SUBAPPLICATION Uebung_157 (* Übung zu FsInfo/FsDir: File Server abfragen und Verzeichnis listen *)
  (* Standard: 61499-2; Description: Copyright (c) 2026 Meisterschulen am Ostbahnhof This program and the accompanying materials are made available under the terms of the Eclipse Public License 2.0 which is available at https://www.eclipse.org/legal/epl-2.0/ SPDX-License-Identifier: EPL-2.0 *)
  (* Version 1.0, 2026-11-26, Franz Höpfinger, Meisterschulen am Ostbahnhof, initial API and implementation and/or initial documentation *)
  PACKAGE Uebungen;
  IMPORT Uebungen::const::Uebung_150_159::FileServer::FS_ADD;
  IMPORT Uebungen::const::Uebung_150_159::FileServer::FS_FLT;
  IMPORT Uebungen::const::Uebung_150_159::FileServer::FS_WURZEL;
  IMPORT isobus::pgn::ISOUSERHOME_e::network;
  IMPORT isobus::pgn::ISO_CAN_NODE::NODE1;
  IMPORT logiBUS::io::DI::logiBUS_DI::Input_I1;
  IMPORT logiBUS::io::DI::logiBUS_DI_Events::BUTTON_SINGLE_CLICK;
  IMPORT logiBUS::io::DQ::logiBUS_DO::Output_Q1;
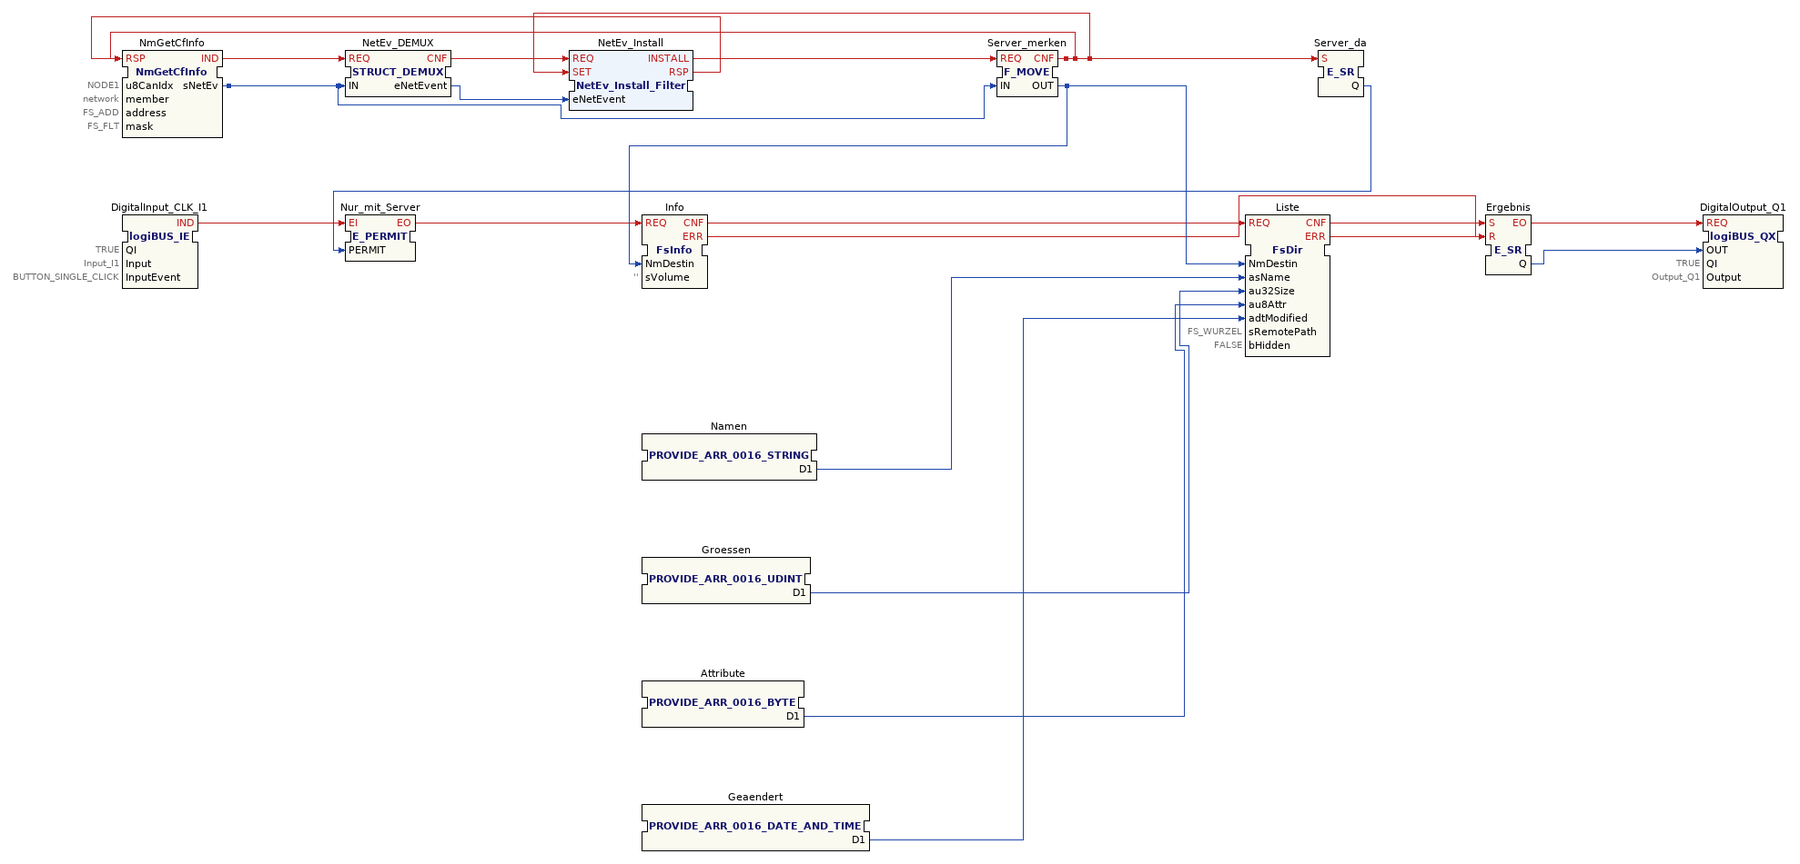
  (* File Server: Eigenschaften abfragen und Verzeichnis listen (FsInfo, FsDir) NmGetCfInfo (network, Filter FS_ADD/FS_FLT = NAME-Funktion 61) meldet den File Server, z. B. CCI 1200 mit USB-Stick. I1 Klick (nur mit Server): FsInfo, dann FsDir auf FS_WURZEL ('.'). Q1 an = fertig, Q1 aus = Fehler. Watch Info: u8Version, u8VolumeStatus (255 = meldet keinen), u32TotalKB, u32FreeKB. Watch Liste: u16Count, asName, au32Size (logibus_test.txt aus Übung 156: 24 Byte). Bei ERR s16Status und u16FsError. Mehr als 16 Einträge: ERR mit E_OVERFLOW (-6), die ersten 16 stehen trotzdem drin. Voraussetzungen: Firmware mit FsInfo/FsDir (neue Host-Symbole), neue isobus_fs-ELF, PART_13_FSC = 1 in /data/functionalities.ini. *)
  FBS
    NmGetCfInfo : isobus::pgn::NmGetCfInfo(u8CanIdx := NODE1, member := network, address := FS_ADD, mask := FS_FLT); (* meldet den File Server (Funktion 61) *)
    NetEv_DEMUX : eclipse4diac::convert::STRUCT_DEMUX; {SET_ATTRIBUTE(StructuredType, isobus::pgn::ISONETEVENT_T)}
    Server_merken : iec61131::selection::F_MOVE; (* eigener CF und File-Server-CF (NmDestin) *)
    Server_da : iec61499::events::E_SR;
    DigitalInput_CLK_I1 : logiBUS::io::DI::logiBUS_IE(QI := TRUE, Input := Input_I1, InputEvent := BUTTON_SINGLE_CLICK);
    Nur_mit_Server : iec61499::events::E_PERMIT;
    Info : isobus::fs::FsInfo(sVolume := ''); (* Version, Volume-Status, Größe und freier Platz *)
    Namen : eclipse4diac::convert::providers::PROVIDE_ARR_0016_STRING;
    Groessen : eclipse4diac::convert::providers::PROVIDE_ARR_0016_UDINT;
    Attribute : eclipse4diac::convert::providers::PROVIDE_ARR_0016_BYTE;
    Geaendert : eclipse4diac::convert::providers::PROVIDE_ARR_0016_DATE_AND_TIME;
    Liste : isobus::fs::FsDir(sRemotePath := FS_WURZEL, bHidden := FALSE); (* Wurzel des aktuellen Volumes, max. 16 Einträge *)
    Ergebnis : iec61499::events::E_SR; (* Q1 an = Info und Liste gelesen *)
    DigitalOutput_Q1 : logiBUS::io::DQ::logiBUS_QX(QI := TRUE, Output := Output_Q1);
  END_FBS
  SUBAPPS
    NetEv_Install : MyLib::sys::NetEv_Install_Filter;
  END_SUBAPPS
  EVENT_CONNECTIONS
    NmGetCfInfo.IND TO NetEv_DEMUX.REQ;
    NetEv_DEMUX.CNF TO NetEv_Install.REQ;
    NetEv_Install.INSTALL TO Server_merken.REQ;
    NetEv_Install.RSP TO NmGetCfInfo.RSP;
    Server_merken.CNF TO NetEv_Install.SET;
    Server_merken.CNF TO Server_da.S;
    Server_merken.CNF TO NmGetCfInfo.RSP;
    DigitalInput_CLK_I1.IND TO Nur_mit_Server.EI;
    Nur_mit_Server.EO TO Info.REQ;
    Info.CNF TO Liste.REQ;
    Liste.CNF TO Ergebnis.S;
    Info.ERR TO Ergebnis.R;
    Liste.ERR TO Ergebnis.R;
    Ergebnis.EO TO DigitalOutput_Q1.REQ;
  END_CONNECTIONS
  DATA_CONNECTIONS
    NmGetCfInfo.sNetEv TO NetEv_DEMUX.IN;
    NetEv_DEMUX.eNetEvent TO NetEv_Install.eNetEvent;
    NmGetCfInfo.sNetEv TO Server_merken.IN;
    Server_merken.OUT TO Info.NmDestin;
    Server_merken.OUT TO Liste.NmDestin;
    Namen.D1 TO Liste.asName;
    Groessen.D1 TO Liste.au32Size;
    Attribute.D1 TO Liste.au8Attr;
    Geaendert.D1 TO Liste.adtModified;
    Server_da.Q TO Nur_mit_Server.PERMIT;
    Ergebnis.Q TO DigitalOutput_Q1.OUT;
  END_CONNECTIONS
END_SUBAPPLICATION
